Universal Robots URScript: T007_mistralai_Mistral-Large-3-675B-Instruct-2512-NVFP4_edit_perf_rep1.urscript

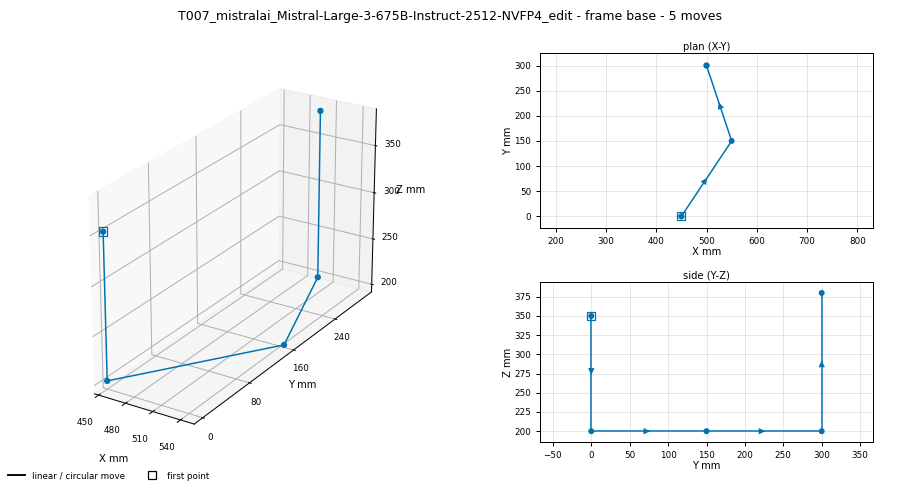
[picture p0: tool path of T007_mistralai_Mistral-Large-3-675B-Instruct-2512-NVFP4_edit_perf_rep1.urscript in frame base, 5 of 7 moves have a stored position in this frame; points joined in program order, loops and branches not executed]
# Task: T007 — Curved contour weld — hybrid mode (optimized)
# Operating mode: hybrid | Max TCP speed: 0.300 m/s
# Robot: ur5e

def task_T007():
  # [0] Verify E-Stop clear
  if (get_digital_in(0) == True):
    popup("E-Stop active — aborting program.", error=True)
    halt
  end

  # [1] Home position - increased acceleration
  movej([0.0000, -1.5708, 1.5708, -1.5708, -1.5708, 0.0000], a=3.0000, v=1.2000)

  # [2] Approach above weld fixture - increased speed and acceleration
  movel(p[0.450000, 0.000000, 0.350000, 0.0000, 3.1416, 0.0000], a=2.0000, v=0.5000, r=0.0100)

  # [3] Descend to weld start - increased acceleration
  movel(p[0.450000, 0.000000, 0.200000, 0.0000, 3.1416, 0.0000], a=1.0000, v=0.1500, r=0.0010)

  # [4] Gas pre-flow ON - parallel with motion
  set_digital_out(1, True)

  # [5] Gas stabilization - reduced time
  sleep(0.3000)

  # [6] Arc ON - parallel with motion start
  set_digital_out(0, True)
  set_analog_out(0, 0.500)
  set_analog_out(1, 0.400)

  # [7] Weld midpoint - increased speed
  movel(p[0.550000, 0.150000, 0.200000, 0.0000, 3.1416, 0.0000], a=0.5000, v=0.1000, r=0.0050)

  # [8] Weld end
  movel(p[0.500000, 0.300000, 0.200000, 0.0000, 3.1416, 0.0000], a=0.5000, v=0.1000)

  # [9] Arc OFF - parallel with motion start
  set_digital_out(0, False)
  set_analog_out(0, 0.0)
  set_analog_out(1, 0.0)

  # [10] Post-weld gas flow - reduced time
  sleep(0.5000)

  # [11] Gas flow OFF
  set_digital_out(1, False)

  # [12] Retract above weld end - increased speed and acceleration
  movel(p[0.500000, 0.300000, 0.380000, 0.0000, 3.1416, 0.0000], a=2.0000, v=0.5000, r=0.0100)

  # [13] Return to home - increased acceleration
  movej([0.0000, -1.5708, 1.5708, -1.5708, -1.5708, 0.0000], a=3.0000, v=1.2000)

end

# Entry point
task_T007()
